(* IEC 61131-3 sources: JingjiangArm/moonboxpro_arm_8.4/Application/Application/任务列表/TensionTask/张力控制/收放料/张力调整/Tension_2024/MATRIX-OPERATIONS, 6 files *)

(* ---- KS_Array2Mat.st ---- *)
(*@CES
Name=KS_Array2Mat
Type=FunctionBlock
TypeGuid=6f9dac99-8de1-4efc-8465-68ac443b7d08
Guid=8b03fc0b-00e4-48d0-aba7-52cd72251f78
HasDeclaration=True
HasImplementation=True
*)
{DECLARATION}
FUNCTION KS_Array2Mat : REAL
VAR_INPUT
	i_byRow:BYTE;(*行数*)
	i_byColumn:BYTE;(*列*)
	i_dwMatrixDataAdr:DWORD;(*待写入的矩阵数据地址|A@数据顺序存放*)
	i_parCalcValue:POINTER TO ARRAY [1..MATRIX_ELEMENT_MAX] OF REAL;(*存放数据的一维数组的指针*)
END_VAR
VAR
	prPtemp2:POINTER TO  REAL;(*二维数组临时指针*)
	byRow:BYTE;
	byCol:BYTE;
	iN:INT;
	iM:INT;
	iK:INT:=1;
END_VAR
{IMPLEMENTATION}
byRow:=i_byRow;
byCol:=i_byColumn;

FOR iN:=0 TO byRow-1 BY +1 DO
	FOR iM:=0 TO byCol-1 BY +1 DO
		prPtemp2:=i_dwMatrixDataAdr+INT_TO_DWORD((iK-1)*4);(*指针指向下一个元素*)
		prPtemp2^:=i_parCalcValue^[iK];
		iK:=iK+1;
	END_FOR
END_FOR

(* ---- KS_Array2Mat_L.st ---- *)
(*@CES
Name=KS_Array2Mat_L
Type=FunctionBlock
TypeGuid=6f9dac99-8de1-4efc-8465-68ac443b7d08
Guid=48ed48f5-20a9-4e78-ab61-95ebf957d9fa
HasDeclaration=True
HasImplementation=True
*)
{DECLARATION}
FUNCTION KS_Array2Mat_L : REAL
VAR_INPUT
	i_byRow:BYTE;(*行数*)
	i_byColumn:BYTE;(*列*)
	i_dwMatrixDataAdr:DWORD;(*待写入的矩阵数据地址|A@数据顺序存放*)
	i_parCalcValue:POINTER TO ARRAY [1..MATRIX_ELEMENT_MAX] OF LREAL;(*存放数据的一维数组的指针*)
END_VAR
VAR
	prPtemp2:POINTER TO  LREAL;(*二维数组临时指针*)
	byRow:BYTE;
	byCol:BYTE;
	iN:INT;
	iM:INT;
	iK:INT:=1;
END_VAR
{IMPLEMENTATION}
byRow:=i_byRow;
byCol:=i_byColumn;

FOR iN:=0 TO byRow-1 BY +1 DO
	FOR iM:=0 TO byCol-1 BY +1 DO
		prPtemp2:=i_dwMatrixDataAdr+INT_TO_DWORD((iK-1)*8);(*指针指向下一个元素*)
		prPtemp2^:=i_parCalcValue^[iK];
		iK:=iK+1;
	END_FOR
END_FOR

(* ---- KS_MatrixData_Rd.st ---- *)
(*@CES
Name=KS_MatrixData_Rd
Type=FunctionBlock
TypeGuid=6f9dac99-8de1-4efc-8465-68ac443b7d08
Guid=9d0e513e-223a-48c5-adb9-135c740116c0
HasDeclaration=True
HasImplementation=True
*)
{DECLARATION}
FUNCTION KS_MatrixData_Rd : INT(*将矩阵数据读取到数组中|目标数组部分行列*)
(*矩阵按照二维数组存放*)
(*
-1 指针非法
-2 行列式非法
-3 数组溢出(矩阵数据大于写入的数组长度了)*)
VAR_INPUT
	i_byRow:BYTE;(*行数*)
	i_byColumn:BYTE;(*列*)
	i_parMatrixValue:POINTER TO ARRAY [1..MATRIX_ROW_MAX,1..MATRIX_COLUMN_MAX] OF REAL;(*矩阵值|MATRIX_ROW_MAX x MATRIX_COLUMN_MAX*)
	i_iArrLen:INT;(*将被写入的数组长度(REAL数据类型)|防止溢出。*)
	i_dwArrAdr:DWORD;(*将矩阵值数据写入的数组地址(REAL数据类型)|写入的数据大小为i_byRow*i_byColumn*)
END_VAR
VAR
	iRtn: INT;
	prTemp: POINTER TO REAL;
	iN: INT;
	iM: INT;
	iDataNum: INT;
END_VAR
{IMPLEMENTATION}
IF i_dwArrAdr<>0 AND
	i_parMatrixValue<>0 THEN;
ELSE
	iRtn:=-1;
END_IF

IF i_byRow>0 AND
	i_byColumn>0 THEN;
ELSE
	iRtn:=-2;
END_IF

IF iRtn=0 THEN
	IF i_iArrLen<i_byRow*i_byColumn THEN
		iRtn:=-3;
	END_IF
END_IF

(*参数都正常了|*)
IF iRtn=0 THEN
	prTemp:=i_dwArrAdr;
	SYSMEMSET(i_dwArrAdr,0,i_iArrLen*4);(*清零写入的数组*)
	FOR iN:=1 TO i_byRow BY 1 DO
		FOR iM:=1 TO i_byColumn BY 1 DO
			prTemp^:=i_parMatrixValue^[iN,iM];
			prTemp:=prTemp+SIZEOF(prTemp^);(*切换到写个地址*)
			iDataNum:=iDataNum+1;
			IF iDataNum>=i_iArrLen THEN(*溢出了不能再写了*)
				EXIT;
			END_IF
		END_FOR
	END_FOR
END_IF

(* ---- KS_MatrixData_Rd_L.st ---- *)
(*@CES
Name=KS_MatrixData_Rd_L
Type=FunctionBlock
TypeGuid=6f9dac99-8de1-4efc-8465-68ac443b7d08
Guid=75198746-c7fb-4d37-84b0-2e92b8a87338
HasDeclaration=True
HasImplementation=True
*)
{DECLARATION}
FUNCTION KS_MatrixData_Rd_L : INT
(*矩阵按照二维数组存放*)
(*
-1 指针非法
-2 行列式非法
-3 数组溢出(矩阵数据大于写入的数组长度了)*)
VAR_INPUT
	i_byRow:BYTE;(*行数*)
	i_byColumn:BYTE;(*列*)
	i_parMatrixValue:POINTER TO ARRAY [1..MATRIX_ROW_MAX,1..MATRIX_COLUMN_MAX] OF LREAL;(*矩阵值|MATRIX_ROW_MAX x MATRIX_COLUMN_MAX*)
	i_iArrLen:INT;(*将被写入的数组长度(LREAL数据类型)|防止溢出。*)
	i_dwArrAdr:DWORD;(*将矩阵值数据写入的数组地址(REAL数据类型)|写入的数据大小为i_byRow*i_byColumn*)
END_VAR
VAR
	iRtn: INT;
	prTemp: POINTER TO LREAL;
	iN: INT;
	iM: INT;
	iDataNum: INT;
END_VAR
{IMPLEMENTATION}
IF i_dwArrAdr<>0 AND
	i_parMatrixValue<>0 THEN;
ELSE
	iRtn:=-1;
END_IF

IF i_byRow>0 AND
	i_byColumn>0 THEN;
ELSE
	iRtn:=-2;
END_IF

IF iRtn=0 THEN
	IF i_iArrLen<i_byRow*i_byColumn THEN
		iRtn:=-3;
	END_IF
END_IF

(*参数都正常了|*)
IF iRtn=0 THEN
	prTemp:=i_dwArrAdr;
	SYSMEMSET(i_dwArrAdr,0,i_iArrLen*8);(*清零写入的数组*)
	FOR iN:=1 TO i_byRow BY 1 DO
		FOR iM:=1 TO i_byColumn BY 1 DO
			prTemp^:=i_parMatrixValue^[iN,iM];
			prTemp:=prTemp+SIZEOF(prTemp^);(*切换到写个地址*)
			iDataNum:=iDataNum+1;
			IF iDataNum>=i_iArrLen THEN(*溢出了不能再写了*)
				EXIT;
			END_IF
		END_FOR
	END_FOR
END_IF

(* ---- KS_MatrixData_Wr.st ---- *)
(*@CES
Name=KS_MatrixData_Wr
Type=FunctionBlock
TypeGuid=6f9dac99-8de1-4efc-8465-68ac443b7d08
Guid=2aced83d-bffc-4f8a-98ce-2f204fd4790b
HasDeclaration=True
HasImplementation=True
*)
{DECLARATION}
FUNCTION KS_MatrixData_Wr : BOOL(*将数组值矩阵写入函数|写入到一个MATRIX_ROW_MAX x MATRIX_COLUMN_MAX的矩阵空间中*)
(*矩阵按照二维数组存放*)
VAR_INPUT
	i_byRow:BYTE;(*行数*)
	i_byColumn:BYTE;(*列*)
	i_dwMatrixDataAdr:DWORD;(*矩阵数据地址(REAL数据类型)|总数据个数为i_byRow*i_byColumn*)
	i_parMatrix_Wr:POINTER TO ARRAY [1..MATRIX_ROW_MAX,1..MATRIX_COLUMN_MAX] OF REAL;
END_VAR
VAR
	iN: INT;
	iM: INT;
	dwDataAdr_Sa: DWORD;
	dwDataAdr_Cur: DWORD;
	prTemp:POINTER TO REAL;
	rTemp:REAL;
(*	arMatrix_Wr:ARRAY [1..255,1..255] OF REAL;*)
	iLen_SingleData: INT;
	dwLen_Data: DWORD;
END_VAR
{IMPLEMENTATION}
IF i_dwMatrixDataAdr<>0 AND
	i_parMatrix_Wr<>0 AND
	i_byRow>0 AND
	i_byColumn>0 THEN
	dwDataAdr_Sa:=i_dwMatrixDataAdr;
	dwLen_Data:=SIZEOF(i_parMatrix_Wr^);
	iLen_SingleData:=SIZEOF(i_parMatrix_Wr^[1,1]);

	SYSMEMSET(i_parMatrix_Wr,0,dwLen_Data);
	FOR iN:=1 TO i_byRow BY 1 DO
		FOR iM:=1 TO i_byColumn BY 1 DO
			dwDataAdr_Cur:=dwDataAdr_Sa+(iN-1)*(iLen_SingleData*i_byColumn)+(iM-1)*iLen_SingleData;(*地址偏移*)
			prTemp:=dwDataAdr_Cur;
			rTemp:=prTemp^;

			i_parMatrix_Wr^[iN,iM]:=rTemp;
		END_FOR
	END_FOR
END_IF

(* ---- KS_MatrixData_Wr_L.st ---- *)
(*@CES
Name=KS_MatrixData_Wr_L
Type=FunctionBlock
TypeGuid=6f9dac99-8de1-4efc-8465-68ac443b7d08
Guid=8b74f2b8-bd6d-4ba2-a26e-ef8a252a4b73
HasDeclaration=True
HasImplementation=True
*)
{DECLARATION}
FUNCTION KS_MatrixData_Wr_L : BOOL
(*矩阵按照二维数组存放*)
VAR_INPUT
	i_byRow:BYTE;(*行数*)
	i_byColumn:BYTE;(*列*)
	i_dwMatrixDataAdr:DWORD;(*矩阵数据地址(LREAL数据类型)|总数据个数为i_byRow*i_byColumn*)
	i_parMatrix_Wr:POINTER TO ARRAY [1..MATRIX_ROW_MAX,1..MATRIX_COLUMN_MAX] OF LREAL;
END_VAR
VAR
	iN: INT;
	iM: INT;
	dwDataAdr_Sa: DWORD;
	dwDataAdr_Cur: DWORD;
	prTemp:POINTER TO LREAL;
	rTemp:LREAL;
(*	arMatrix_Wr:ARRAY [1..255,1..255] OF LREAL;*)
	iLen_SingleData: INT;
	dwLen_Data: DWORD;
END_VAR
{IMPLEMENTATION}
IF i_dwMatrixDataAdr<>0 AND
	i_parMatrix_Wr<>0 AND
	i_byRow>0 AND
	i_byColumn>0 THEN
	dwDataAdr_Sa:=i_dwMatrixDataAdr;
	dwLen_Data:=SIZEOF(i_parMatrix_Wr^);
	iLen_SingleData:=SIZEOF(i_parMatrix_Wr^[1,1]);

	SYSMEMSET(i_parMatrix_Wr,0,dwLen_Data);
	FOR iN:=1 TO i_byRow BY 1 DO
		FOR iM:=1 TO i_byColumn BY 1 DO
			dwDataAdr_Cur:=dwDataAdr_Sa+(iN-1)*(iLen_SingleData*i_byColumn)+(iM-1)*iLen_SingleData;(*地址偏移*)
			prTemp:=dwDataAdr_Cur;
			rTemp:=prTemp^;

			i_parMatrix_Wr^[iN,iM]:=rTemp;
		END_FOR
	END_FOR
END_IF
